// TIA Portal V19 export
TYPE "ST_Error"
   STRUCT
      "Bit:0" : Bool;
      "Bit:1" : Bool;
      "Bit:2" : Bool;
      "Bit:3" : Bool;
      "Bit:4" : Bool;
      "Bit:5" : Bool;
      "Bit:6" : Bool;
      "Bit:7" : Bool;
      "Bit:8" : Bool;
      "Bit:9" : Bool;
      "Bit:10" : Bool;
      "Bit:11" : Bool;
      "Bit:12" : Bool;
      "Bit:13" : Bool;
      "Bit:14" : Bool;
      "Bit:15" : Bool;
      "Bit:16" : Bool;
      "Bit:17" : Bool;
      "Bit:18" : Bool;
      "Bit:19" : Bool;
      "Bit:20" : Bool;
      "Bit:21" : Bool;
      "Bit:22" : Bool;
      "Bit:23" : Bool;
      "Bit:24" : Bool;
      "Bit:25" : Bool;
      "Bit:26" : Bool;
      "Bit:27" : Bool;
      "Bit:28" : Bool;
      "Bit:29" : Bool;
      "Bit:30" : Bool;
      "Bit:31" : Bool;
      "Bit:32" : Bool;
   END_STRUCT;
END_TYPE
